          Waypoint Variable (Variable): motionParameters(jointSpeed=1.047198 jointAcceleration=1.396263 cartesianSpeed=0.09 cartesianAcceleration=0.05); variable=PSE_T_H
          URCap Gripper (Robotiq_Grippers, Robotiq Inc.) dataModel(position=24.705882352941178, force=11.0, speed=0.0, positionInDouble=24.705882352941178, forceInDouble=11.0, speedInDouble=0.0, slaveIds=[9], blocking=true)
          Waypoint Variable (Variable): variable=PSE_R
    Case (caseValue=7)
      Folder Load [hidden by the author, left out]
    Case (caseValue=8)
      Folder Unload [hidden by the author, left out]
    Case (caseValue=11)
      Folder Place without opening gripper
        Action_Info := "place object without gripper opening"
        Script: do_transition(pose_trans(FRM_Reference, PSE_T), keep_rxry=OBJ_Picked)
        Folder EXTT
          Switch expression=JIG
            Case (caseValue=1)
              Folder 3FG
                If OBJ_Picked
                  Set DigitalOutput pin=GRP_3F_Open; digitalValue=1
        If PSE_A_H≠PSE_Z
          If JNT_Q≠JNT_Z
            Script: movej(get_inverse_kin(pose_trans(FRM_Reference, PSE_A_H), qnear=JNT_Q), r=0.050)
          Else 
            Script: movej(pose_trans(FRM_Reference, PSE_A_H), r=0.050)
        If PSE_A≠PSE_Z
          If JNT_Q≠JNT_Z
            Script: movej(get_inverse_kin(pose_trans(FRM_Reference, PSE_A), qnear=JNT_Q), r=0.020)
          Else 
            Script: movej(pose_trans(FRM_Reference, PSE_A), r=0.020)
        MoveL speed 400 mm/s, acceleration 500 mm/s^2 (useActiveTCP=true) feature=FRM_Reference
          If PSE_T_H≠PSE_Z
            Waypoint Variable (Variable): motionParameters(blendRadius=0.01); variable=PSE_T_H
          Waypoint Variable (Variable): motionParameters(jointSpeed=1.047198 jointAcceleration=1.396263 cartesianSpeed=0.09 cartesianAcceleration=0.05); variable=PSE_T
            Until TOOL_CONTACT_DETECTION (allowActions=false retraction=NONE decelerationAcceleration=0.5 decelerationAngularAcceleration=34.906585)
          Force Frame feature=FRM_Reference; selection=[1, 1, 1, 0, 0, 0]; wrench=[0, 0, 0, 0, 0, 0]; limitsForce=[0.1, 0.1, 0.01, 1.047198, 1.047198, 1.047198]; limitsMotion=[0.1, 0.1, 0.1, 0.349066, 0.349066, 0.349066]
            Waypoint Variable (Variable): motionParameters(jointSpeed=1.047198 jointAcceleration=1.396263 cartesianSpeed=0.07 cartesianAcceleration=0.04); variable=PSE_T
          Folder EXTT
            Switch expression=JIG
              Case (caseValue=1)
                Folder 3FG
                  If OBJ_Picked
                    Set DigitalOutput pin=GRP_3F_Open; digitalValue=0
                    Wait Sleep waitTime=0.2
          Folder EOAT
            ''
    Case (caseValue=12)
      Folder Decap
        Action_Info := "decapping"
        Set DigitalOutput pin=GRP_3F_Enable; digitalValue=1
        Set DigitalOutput pin=GRP_3F_Decap; digitalValue=1
        Force Simple feature=Joint_6_name; selection=[0, 0, 1, 0, 0, 0]; wrench=[0, 0, 5, 0, 0, 0]; limitsForce=[0.15, 0.15, 0.15, 1.047198, 1.047198, 1.047198]; limitsMotion=[0.1, 0.1, 0.1, 0.349066, 0.349066, 0.349066]
          Script: check_decapping(offset=0.015, timeout=5, abort=CMD_Hold)
        Set DigitalOutput pin=GRP_3F_Decap; digitalValue=0
        Set DigitalOutput pin=GRP_3F_Enable; digitalValue=0
        MoveL speed 150 mm/s, acceleration 800 mm/s^2 (useActiveTCP=true) feature=FRM_Reference
          Waypoint Variable (Variable): variable=PSE_R
    Case (caseValue=13)
      Timer (action=Reset) variable(name=TMR_Barcode)
      Folder Read [hidden by the author, left out]
    Case (caseValue=15)
      Folder Detect
        Action_Info := "detect"
    Case (caseValue=30)
      Folder Shake
        Action_Info := "shake"
        Script: do_transition(pose_trans(FRM_Reference, PSE_T), keep_rxry=OBJ_Picked)
        If PSE_A_H≠PSE_Z
          If JNT_Q≠JNT_Z
            Script: movej(get_inverse_kin(pose_trans(FRM_Reference, PSE_A_H), qnear=JNT_Q), r=0.050)
          Else 
            Script: movej(pose_trans(FRM_Reference, PSE_A_H), r=0.050)
        If PSE_A≠PSE_Z
          If JNT_Q≠JNT_Z
            Script: movej(get_inverse_kin(pose_trans(FRM_Reference, PSE_A), qnear=JNT_Q), r=0.020)
          Else 
            Script: movej(pose_trans(FRM_Reference, PSE_A), r=0.020)
        MoveL speed 400 mm/s, acceleration 500 mm/s^2 (useActiveTCP=true) feature=FRM_Reference
          If PSE_T_H≠PSE_Z
            Waypoint Variable (Variable): motionParameters(blendRadius=0.01); variable=PSE_T_H
          Waypoint Variable (Variable): motionParameters(jointSpeed=1.047198 jointAcceleration=1.396263 cartesianSpeed=0.12 cartesianAcceleration=0.08); variable=PSE_T
          Folder EXTT
            ''
            MoveJ speed 60 deg/s, acceleration 80 deg/s^2 (useActiveTCP=true) feature=Base
              Waypoint Waypoint_6: TCP in base x=8.801 y=-547.927 z=402.697 mm, rx=-0.5899 ry=-0.0072 rz=-0.0613 rad; joints [-69.01, -76.872, -104.694, -56.634, 78.043, -158.781] deg; TCP offset x=0 y=0 z=161 mm, rx=3.1415 ry=0 rz=0 rad
            MoveJ speed 60 deg/s, acceleration 80 deg/s^2 (useActiveTCP=true) feature=Base
              Waypoint Waypoint_18: TCP in base x=-178.372 y=-433.927 z=368.082 mm, rx=-0.0866 ry=0.7047 rz=-0.0079 rad; joints [-72.502, -76.524, -102.817, -99.71, 50.308, -158.785] deg
            MoveJ speed 60 deg/s, acceleration 80 deg/s^2 (useActiveTCP=true) feature=Base
              Waypoint Waypoint_12: TCP in base x=8.801 y=-547.927 z=402.697 mm, rx=-0.5899 ry=-0.0072 rz=-0.0613 rad; joints [-69.01, -76.872, -104.694, -56.634, 78.043, -158.781] deg
            MoveJ speed 60 deg/s, acceleration 80 deg/s^2 (useActiveTCP=true) feature=Base
              Waypoint Waypoint_19: TCP in base x=-178.372 y=-433.927 z=368.082 mm, rx=-0.0866 ry=0.7047 rz=-0.0079 rad; joints [-72.502, -76.524, -102.817, -99.71, 50.308, -158.785] deg
          If PSE_R_H≠PSE_Z
            Waypoint Variable (Variable): motionParameters(blendRadius=0.01); variable=PSE_R
            Waypoint Variable (Variable): variable=PSE_R_H
          Else 
            Waypoint Variable (Variable): variable=PSE_R
    Case (caseValue=31)
      Action_Info := "Pick_Vial"
      Folder Pick_Vial
        URCap Gripper (Robotiq_Grippers, Robotiq Inc.) dataModel(position=0.0, force=27.84313725490196, speed=32.15686274509804, positionInDouble=0.0, forceInDouble=27.84313725490196, speedInDouble=32.15686274509804, slaveIds=[9], blocking=true)
        MoveJ speed 60 deg/s, acceleration 80 deg/s^2 (useActiveTCP=true) feature=Base
          Waypoint Vial_above: motionParameters(jointSpeed=0.436332 jointAcceleration=0.523599 cartesianSpeed=0.25 cartesianAcceleration=1.2 blendRadius=0.05); TCP in base x=17.106 y=-652.093 z=184.921 mm, rx=0 ry=0 rz=1.5641 rad; joints [-76.636, -112.403, -84.029, -73.556, 90.141, -256.27] deg
        MoveL speed 250 mm/s, acceleration 1200 mm/s^2 (useActiveTCP=true) feature=Base
          Waypoint Vial_pick_point: motionParameters(jointSpeed=1.047198 jointAcceleration=1.396263 cartesianSpeed=0.1 cartesianAcceleration=0.5); TCP in base x=17.106 y=-648.923 z=93.308 mm, rx=0 ry=0 rz=1.5641 rad; joints [-76.583, -116.742, -92.083, -61.164, 90.132, -256.177] deg
        URCap Gripper (Robotiq_Grippers, Robotiq Inc.) dataModel(position=100.0, force=32.94117647058823, speed=27.84313725490196, positionInDouble=100.0, forceInDouble=32.94117647058823, speedInDouble=27.84313725490196, slaveIds=[9], blocking=true)
        MoveL speed 250 mm/s, acceleration 1200 mm/s^2 (useActiveTCP=true) feature=Base
          Waypoint Waypoint_20: motionParameters(jointSpeed=1.047198 jointAcceleration=1.396263 cartesianSpeed=0.1 cartesianAcceleration=0.5 blendRadius=0.05); TCP in base x=19.228 y=-648.67 z=184.921 mm, rx=0 ry=0 rz=0.0241 rad; joints [-76.382, -111.96, -84.66, -73.372, 90.146, -167.779] deg
        SafeHome (positionOptionType=SPEED_AND_ACCELERATION speed=1.047198 acceleration=1.396263 nextMotionTime=2)
    Case (caseValue=32)
      decap := False
      Folder decap_Vial
        Set DigitalOutput pin=digital_out[5]; digitalValue=1
        MoveJ speed 60 deg/s, acceleration 80 deg/s^2 (useActiveTCP=true) feature=Base
          Waypoint Waypoint_47: motionParameters(jointSpeed=0.436332 jointAcceleration=0.523599 cartesianSpeed=0.25 cartesianAcceleration=1.2 blendRadius=0); TCP in base x=-32.362 y=-348.336 z=391.476 mm, rx=0 ry=0 rz=-0.0047 rad; joints [-72.819, -68.266, -97.918, -103.808, 90.124, -162.602] deg
        MoveL speed 250 mm/s, acceleration 1200 mm/s^2 (useActiveTCP=true) feature=Base
          Waypoint Vial_3FG_place: motionParameters(jointSpeed=1.047198 jointAcceleration=1.396263 cartesianSpeed=0.1 cartesianAcceleration=0.5); TCP in base x=-31.859 y=-349.403 z=145.301 mm, rx=0 ry=0 rz=0 rad; joints [-72.903, -71.756, -132.514, -65.722, 90.129, -162.805] deg
        Set DigitalOutput pin=digital_out[5]; digitalValue=0
        Wait Sleep waitTime=0.5
        MoveL speed 250 mm/s, acceleration 1200 mm/s^2 (useActiveTCP=true) feature=Base
          Waypoint Waypoint_48: motionParameters(jointSpeed=1.047198 jointAcceleration=1.396263 cartesianSpeed=0.1 cartesianAcceleration=0.5 blendRadius=0.05); TCP in base x=-32.362 y=-348.336 z=391.476 mm, rx=0 ry=0 rz=-0.0047 rad; joints [-72.819, -68.266, -97.918, -103.808, 90.124, -162.602] deg
        MoveJ speed 60 deg/s, acceleration 80 deg/s^2 (useActiveTCP=true) feature=Base
          Waypoint cap_dump: motionParameters(jointSpeed=0.436332 jointAcceleration=0.523599 cartesianSpeed=0.25 cartesianAcceleration=1.2); TCP in base x=-139.169 y=-420.164 z=146.096 mm, rx=0 ry=0 rz=0 rad; joints [-90.79, -86.479, -121, -62.513, 90.12, -180.712] deg
        URCap Gripper (Robotiq_Grippers, Robotiq Inc.) dataModel(position=0.0, force=100.0, speed=100.0, positionInDouble=0.0, forceInDouble=100.0, speedInDouble=100.0, slaveIds=[9], blocking=true)
        MoveJ speed 60 deg/s, acceleration 80 deg/s^2 (useActiveTCP=true) feature=Base
          Waypoint Waypoint_49: motionParameters(jointSpeed=0.436332 jointAcceleration=0.523599 cartesianSpeed=0.25 cartesianAcceleration=1.2 blendRadius=0.05); TCP in base x=-32.362 y=-348.336 z=391.476 mm, rx=0 ry=0 rz=-0.0047 rad; joints [-72.819, -68.266, -97.918, -103.808, 90.124, -162.602] deg
        MoveL speed 250 mm/s, acceleration 1200 mm/s^2 (useActiveTCP=true) feature=Base
          Waypoint Vial_3FG_place: motionParameters(jointSpeed=1.047198 jointAcceleration=1.396263 cartesianSpeed=0.1 cartesianAcceleration=0.5); TCP in base x=-31.859 y=-349.403 z=145.301 mm, rx=0 ry=0 rz=0 rad; joints [-72.903, -71.756, -132.514, -65.722, 90.129, -162.805] deg
        URCap Gripper (Robotiq_Grippers, Robotiq Inc.) dataModel(position=100.0, force=100.0, speed=80.0, positionInDouble=100.0, forceInDouble=100.0, speedInDouble=80.0, slaveIds=[9], blocking=true)
        SuppressedNode
          decap := True
        SuppressedNode
          Script: dynamic_upward_motion(0.015, 7)
        SuppressedNode
          MoveL speed 250 mm/s, acceleration 1200 mm/s^2 (useActiveTCP=true) feature=Joint_6_name
            MoveDirectionNode (selectedDirection=ZPlus toolParams=8.0E-4, 0.001) feature=Base
              Until DISTANCE (allowActions=false deceleration=3 distanceNodeType=STOP) Distance=0.01; motionParameters(blendRadius=0)
        SuppressedNode
          decap := False
        Folder Decap
          Action_Info := "decapping"
          Set DigitalOutput pin=GRP_3F_Enable; digitalValue=1
          Set DigitalOutput pin=GRP_3F_Decap; digitalValue=1
          Force Frame feature=Base; selection=[0, 0, 1, 0, 0, 0]; wrench=[0, 0, 1, 0, 0, 0]; limitsForce=[0.15, 0.15, 0.001, 1.047198, 1.047198, 1.047198]; limitsMotion=[0.1, 0.1, 0.1, 0.349066, 0.349066, 0.349066]
            Script: check_decapping(offset=0.015, timeout=10, abort=CMD_Hold)
          Set DigitalOutput pin=GRP_3F_Decap; digitalValue=0
          Set DigitalOutput pin=GRP_3F_Enable; digitalValue=0
          MoveL speed 250 mm/s, acceleration 1200 mm/s^2 (useActiveTCP=true) feature=Base
            Waypoint Waypoint_50: motionParameters(jointSpeed=1.047198 jointAcceleration=1.396263 cartesianSpeed=0.1 cartesianAcceleration=0.5 blendRadius=0.05); TCP in base x=-32.362 y=-348.336 z=391.476 mm, rx=0 ry=0 rz=-0.0047 rad; joints [-72.819, -68.266, -97.918, -103.808, 90.124, -162.602] deg
        MoveJ speed 60 deg/s, acceleration 80 deg/s^2 (useActiveTCP=true) feature=Base
          Waypoint cap_dump: motionParameters(jointSpeed=0.436332 jointAcceleration=0.523599 cartesianSpeed=0.25 cartesianAcceleration=1.2); TCP in base x=-139.169 y=-420.164 z=146.096 mm, rx=0 ry=0 rz=0 rad; joints [-90.79, -86.479, -121, -62.513, 90.12, -180.712] deg
        URCap Gripper (Robotiq_Grippers, Robotiq Inc.) dataModel(position=0.0, force=100.0, speed=80.0, positionInDouble=0.0, forceInDouble=100.0, speedInDouble=80.0, slaveIds=[9], blocking=true)
        MoveJ speed 60 deg/s, acceleration 80 deg/s^2 (useActiveTCP=true) feature=Base
          Waypoint Waypoint_51: motionParameters(jointSpeed=0.436332 jointAcceleration=0.523599 cartesianSpeed=0.25 cartesianAcceleration=1.2 blendRadius=0.036); TCP in base x=-32.362 y=-348.336 z=391.476 mm, rx=0 ry=0 rz=-0.0047 rad; joints [-72.819, -68.266, -97.918, -103.808, 90.124, -162.602] deg
    Case (caseValue=33)
      Folder Shake and liquid transfer
        MoveL speed 250 mm/s, acceleration 1200 mm/s^2 (useActiveTCP=true) feature=Base
          Waypoint Vial_liq_above: motionParameters(jointSpeed=1.047198 jointAcceleration=1.396263 cartesianSpeed=0.1 cartesianAcceleration=0.5); TCP in base x=-25.304 y=-338.759 z=426.628 mm, rx=-1.3159 ry=0.8 rz=-0.9283 rad; joints [-21.713, -86.8, -129.663, 45.096, -43.028, -184.708] deg
          Waypoint Vial_liq_pick_1: motionParameters(jointSpeed=1.047198 jointAcceleration=1.396263 cartesianSpeed=0.1 cartesianAcceleration=0.5); TCP in base x=-2.66 y=-335.985 z=159.39 mm, rx=-1.1505 ry=0.6732 rz=-1.0106 rad; joints [-20.975, -83.1, -137.831, -114.287, 46.064, -14.375] deg
          Waypoint Vial_liq_pick_2: motionParameters(jointSpeed=1.047198 jointAcceleration=1.396263 cartesianSpeed=0.1 cartesianAcceleration=0.5); TCP in base x=-41.402 y=-356.792 z=125.395 mm, rx=-1.1435 ry=0.6511 rz=-0.8787 rad; joints [-25.36, -82.348, -146.215, -101.788, 37.598, -24.648] deg
          URCap Gripper (Robotiq_Grippers, Robotiq Inc.) dataModel(position=100.0, force=27.84313725490196, speed=32.15686274509804, positionInDouble=100.0, forceInDouble=27.84313725490196, speedInDouble=32.15686274509804, slaveIds=[9], blocking=true)
          Wait Sleep waitTime=1
          Set DigitalOutput pin=digital_out[5]; digitalValue=1
          Wait Sleep waitTime=0.5
          Waypoint Vial_liq_above: motionParameters(jointSpeed=1.047198 jointAcceleration=1.396263 cartesianSpeed=0.05 cartesianAcceleration=0.3 blendRadius=0.05); TCP in base x=-25.304 y=-338.759 z=426.628 mm, rx=-1.3159 ry=0.8 rz=-0.9283 rad; joints [-21.713, -86.8, -129.663, 45.096, -43.028, -184.708] deg
        MoveL speed 250 mm/s, acceleration 1200 mm/s^2 (useActiveTCP=true) feature=Base
          Waypoint Liquid_midway: motionParameters(jointSpeed=1.047198 jointAcceleration=1.396263 cartesianSpeed=0.1 cartesianAcceleration=0.5 blendRadius=0); TCP in base x=57.575 y=-583.082 z=306.415 mm, rx=-1.3517 ry=0.1209 rz=-0.0969 rad; joints [-51.29, -97.606, -136.419, 36.185, 44.156, -168.768] deg
          Loop Counting (count=3) loopVariable(name=Loop_1)
            Waypoint shake_1: motionParameters(jointSpeed=1.047198 jointAcceleration=1.396263 cartesianSpeed=0.5 cartesianAcceleration=2); TCP in base x=57.575 y=-583.085 z=306.423 mm, rx=-1.361 ry=-0.1556 rz=-0.4381 rad; joints [-51.29, -97.606, -136.418, 36.185, 44.156, -145.5] deg
            Waypoint shake_2: motionParameters(jointSpeed=1.047198 jointAcceleration=1.396263 cartesianSpeed=0.5 cartesianAcceleration=2); TCP in base x=57.582 y=-583.091 z=306.44 mm, rx=-1.3088 ry=0.3685 rz=0.2149 rad; joints [-51.29, -97.606, -136.416, 36.185, 44.155, -190] deg
          Waypoint drop_above_1: motionParameters(jointSpeed=1.047198 jointAcceleration=1.396263 cartesianSpeed=0.1 cartesianAcceleration=0.5); TCP in base x=268.235 y=-467.784 z=226.22 mm, rx=-1.0278 ry=-0.4308 rz=1.0046 rad; joints [-53.609, -95.474, -138.959, 24.045, 105.829, -198.245] deg
          Waypoint drop_above_2: motionParameters(jointSpeed=1.047198 jointAcceleration=1.396263 cartesianSpeed=0.1 cartesianAcceleration=0.5); TCP in base x=219.042 y=-470.776 z=133.754 mm, rx=-0.313 ry=-0.3444 rz=1.5006 rad; joints [-60.743, -97.429, -119.175, -41.501, 111.324, -235.78] deg
          Waypoint liq_tran_1: motionParameters(jointSpeed=1.047198 jointAcceleration=1.396263 cartesianSpeed=0.05 cartesianAcceleration=0.5 blendRadius=0.008); TCP in base x=213.068 y=-469.567 z=100.231 mm, rx=0.2519 ry=0.2179 rz=1.5928 rad; joints [-44.631, -104.414, -106.819, -71.743, 78.886, -225.335] deg
          Wait Sleep waitTime=1
          Waypoint drop_above_2: motionParameters(jointSpeed=1.047198 jointAcceleration=1.396263 cartesianSpeed=0.1 cartesianAcceleration=0.5); TCP in base x=219.042 y=-470.776 z=133.754 mm, rx=-0.313 ry=-0.3444 rz=1.5006 rad; joints [-60.743, -97.429, -119.175, -41.501, 111.324, -235.78] deg
          Waypoint Waypoint_21: motionParameters(jointSpeed=1.047198 jointAcceleration=1.396263 cartesianSpeed=0.1 cartesianAcceleration=0.5); TCP in base x=187.119 y=-493.959 z=133.754 mm, rx=-0.313 ry=-0.3444 rz=1.5006 rad; joints [-65.422, -99.182, -116.519, -44.234, 112.218, -240.733] deg
          Waypoint liq_tran_2: motionParameters(jointSpeed=1.047198 jointAcceleration=1.396263 cartesianSpeed=0.05 cartesianAcceleration=0.5); TCP in base x=195.958 y=-493.023 z=100.231 mm, rx=0.1607 ry=0.1098 rz=1.5253 rad; joints [-50.52, -104.533, -106.862, -66.514, 83.832, -227.689] deg
          Wait Sleep waitTime=1
          Waypoint drop_above_2: motionParameters(jointSpeed=1.047198 jointAcceleration=1.396263 cartesianSpeed=0.1 cartesianAcceleration=0.5); TCP in base x=219.042 y=-470.776 z=133.754 mm, rx=-0.313 ry=-0.3444 rz=1.5006 rad; joints [-60.743, -97.429, -119.175, -41.501, 111.324, -235.78] deg
          Waypoint drop_above_1: motionParameters(jointSpeed=1.047198 jointAcceleration=1.396263 cartesianSpeed=0.1 cartesianAcceleration=0.5); TCP in base x=268.235 y=-467.784 z=226.22 mm, rx=-1.0278 ry=-0.4308 rz=1.0046 rad; joints [-53.609, -95.474, -138.959, 24.045, 105.829, -198.245] deg
          Waypoint Liquid_midway: motionParameters(jointSpeed=1.047198 jointAcceleration=1.396263 cartesianSpeed=0.1 cartesianAcceleration=0.5); TCP in base x=57.575 y=-583.082 z=306.415 mm, rx=-1.3517 ry=0.1209 rz=-0.0969 rad; joints [-51.29, -97.606, -136.419, 36.185, 44.156, -168.768] deg
        MoveL speed 250 mm/s, acceleration 1200 mm/s^2 (useActiveTCP=true) feature=Base
          Waypoint Vial_drop_above: motionParameters(jointSpeed=1.047198 jointAcceleration=1.396263 cartesianSpeed=0.1 cartesianAcceleration=0.5); TCP in base x=0.325 y=-648.57 z=221.894 mm, rx=-0.8735 ry=1.1659 rz=-1.4827 rad; joints [-60.601, -137.11, -52.92, -147.418, 45.283, -19.072] deg
          Waypoint Vial_liq_drop: motionParameters(jointSpeed=1.047198 jointAcceleration=1.396263 cartesianSpeed=0.1 cartesianAcceleration=0.5); TCP in base x=1.021 y=-647.66 z=92.916 mm, rx=-0.8348 ry=1.0819 rz=-1.5406 rad; joints [-60.917, -140.075, -64.676, -125.954, 46.582, -22.337] deg
          URCap Gripper (Robotiq_Grippers, Robotiq Inc.) dataModel(position=0.0, force=27.84313725490196, speed=32.15686274509804, positionInDouble=0.0, forceInDouble=27.84313725490196, speedInDouble=32.15686274509804, slaveIds=[9], blocking=true)
          Waypoint Vial_drop_above: motionParameters(jointSpeed=1.047198 jointAcceleration=1.396263 cartesianSpeed=0.1 cartesianAcceleration=0.5); TCP in base x=0.325 y=-648.57 z=221.894 mm, rx=-0.8735 ry=1.1659 rz=-1.4827 rad; joints [-60.601, -137.11, -52.92, -147.418, 45.283, -19.072] deg
    Case (caseValue=34)
      SafeHome (positionOptionType=SPEED_AND_ACCELERATION speed=1.047198 acceleration=1.396263 nextMotionTime=2)
      MoveJ speed 60 deg/s, acceleration 80 deg/s^2 (useActiveTCP=true) feature=Base
        Waypoint Waypoint_9: motionParameters(jointSpeed=0.436332 jointAcceleration=0.523599 cartesianSpeed=0.25 cartesianAcceleration=1.2); TCP in base x=206.301 y=-401.796 z=209.941 mm, rx=0 ry=0 rz=1.5608 rad; joints [-45.627, -84.145, -113.025, -72.821, 90.127, -225.014] deg
      MoveL speed 250 mm/s, acceleration 1200 mm/s^2 (useActiveTCP=true) feature=Base
        Waypoint Waypoint_10: motionParameters(jointSpeed=1.047198 jointAcceleration=1.396263 cartesianSpeed=0.1 cartesianAcceleration=0.5); TCP in base x=200.866 y=-400.818 z=105.073 mm, rx=0 ry=0 rz=1.5608 rad; joints [-46.083, -90.669, -123.933, -55.389, 90.105, -225.416] deg
      URCap Gripper (Robotiq_Grippers, Robotiq Inc.) dataModel(position=100.0, force=27.84313725490196, speed=32.15686274509804, positionInDouble=100.0, forceInDouble=27.84313725490196, speedInDouble=32.15686274509804, slaveIds=[9], blocking=true)
      Wait Sleep waitTime=1
      MoveL speed 250 mm/s, acceleration 1200 mm/s^2 (useActiveTCP=true) feature=Base
        Waypoint Waypoint_11: motionParameters(jointSpeed=1.047198 jointAcceleration=1.396263 cartesianSpeed=0.1 cartesianAcceleration=0.5 blendRadius=0.05); TCP in base x=200.866 y=-400.818 z=325.177 mm, rx=0 ry=0 rz=1.5608 rad; joints [-46.018, -81.306, -98.396, -90.289, 90.129, -225.47] deg
      MoveJ speed 60 deg/s, acceleration 80 deg/s^2 (useActiveTCP=true) feature=Base
        Waypoint Waypoint_7: motionParameters(jointSpeed=0.436332 jointAcceleration=0.523599 cartesianSpeed=0.25 cartesianAcceleration=1.2 blendRadius=0.05); TCP in base x=-615.829 y=233.809 z=300 mm, rx=0.0051 ry=0.0087 rz=-2.1118 rad; joints [-188.832, -110.936, -69.076, -89.912, 89.674, -157.919] deg
      MoveL speed 250 mm/s, acceleration 1200 mm/s^2 (useActiveTCP=true) feature=Base
        Waypoint Waypoint_8: motionParameters(jointSpeed=1.047198 jointAcceleration=1.396263 cartesianSpeed=0.1 cartesianAcceleration=0.5); TCP in base x=-615.829 y=233.809 z=13.91 mm, rx=0.0051 ry=0.0087 rz=-2.1118 rad; joints [-188.874, -123.68, -94.539, -51.707, 89.657, -157.833] deg
      URCap Gripper (Robotiq_Grippers, Robotiq Inc.) dataModel(position=0.0, force=27.84313725490196, speed=32.15686274509804, positionInDouble=0.0, forceInDouble=27.84313725490196, speedInDouble=32.15686274509804, slaveIds=[9], blocking=true)
      MoveJ speed 60 deg/s, acceleration 80 deg/s^2 (useActiveTCP=true) feature=Base
        Waypoint Waypoint_7: motionParameters(jointSpeed=0.436332 jointAcceleration=0.523599 cartesianSpeed=0.25 cartesianAcceleration=1.2); TCP in base x=-615.829 y=233.809 z=300 mm, rx=0.0051 ry=0.0087 rz=-2.1118 rad; joints [-188.832, -110.936, -69.076, -89.912, 89.674, -157.919] deg
      SafeHome (positionOptionType=SPEED_AND_ACCELERATION speed=1.047198 acceleration=1.396263 nextMotionTime=2)
      SuppressedNode
        Folder Decap
          Action_Info := "decapping"
          Set DigitalOutput pin=GRP_3F_Enable; digitalValue=1
          Set DigitalOutput pin=GRP_3F_Decap; digitalValue=1
          Force Frame feature=Base; selection=[0, 0, 1, 0, 0, 0]; wrench=[0, 0, 1, 0, 0, 0]; limitsForce=[0.15, 0.15, 0.001, 1.047198, 1.047198, 1.047198]; limitsMotion=[0.1, 0.1, 0.1, 0.349066, 0.349066, 0.349066]
            Script: check_decapping(offset=0.015, timeout=10, abort=CMD_Hold)
          Set DigitalOutput pin=GRP_3F_Decap; digitalValue=0
          Set DigitalOutput pin=GRP_3F_Enable; digitalValue=0
          MoveL speed 250 mm/s, acceleration 1200 mm/s^2 (useActiveTCP=true) feature=Base
            Waypoint Waypoint_5: motionParameters(jointSpeed=1.047198 jointAcceleration=1.396263 cartesianSpeed=0.1 cartesianAcceleration=0.5 blendRadius=0.05); TCP in base x=-31.859 y=-349.402 z=312.809 mm, rx=0 ry=0 rz=0 rad; joints [-72.832, -66.838, -110.376, -92.778, 90.139, -162.834] deg
          MoveJ speed 60 deg/s, acceleration 80 deg/s^2 (useActiveTCP=true) feature=Base
            Waypoint cap_dump: motionParameters(jointSpeed=0.436332 jointAcceleration=0.523599 cartesianSpeed=0.25 cartesianAcceleration=1.2); TCP in base x=-139.169 y=-420.164 z=146.096 mm, rx=0 ry=0 rz=0 rad; joints [-90.79, -86.479, -121, -62.513, 90.12, -180.712] deg
          URCap Gripper (Robotiq_Grippers, Robotiq Inc.) dataModel(position=0.0, force=100.0, speed=100.0, positionInDouble=0.0, forceInDouble=100.0, speedInDouble=100.0, slaveIds=[9], blocking=true)
          MoveJ speed 60 deg/s, acceleration 80 deg/s^2 (useActiveTCP=true) feature=Base
            Waypoint Waypoint_5: motionParameters(jointSpeed=0.436332 jointAcceleration=0.523599 cartesianSpeed=0.25 cartesianAcceleration=1.2 blendRadius=0.05); TCP in base x=-31.859 y=-349.402 z=312.809 mm, rx=0 ry=0 rz=0 rad; joints [-72.832, -66.838, -110.376, -92.778, 90.139, -162.834] deg
          Set DigitalOutput pin=digital_out[5]; digitalValue=1
    Case (caseValue=35)
      Folder Pick the powder container
        Wait Sleep waitTime=1
        MoveJ speed 60 deg/s, acceleration 80 deg/s^2 (useActiveTCP=true) feature=Base
          Waypoint Container_midwa: motionParameters(blendRadius=0.05); TCP in base x=-379.239 y=-127.191 z=300 mm, rx=0 ry=0 rz=-1.2472 rad; joints [-141.945, -74.312, -107.466, -88.214, 90.137, -160.485] deg
          Waypoint Container_capt: TCP in base x=-525.59 y=407.248 z=411.588 mm, rx=0 ry=0 rz=-2.8961 rad; joints [-206.083, -114.879, -46.847, -108.265, 90.132, -130.312] deg
        URCap VISOR Robotic App (SensoPart VISOR Robotic, SensoPart Industriesensorik GmbH) dataModel(visorAppTemplate=1); state(isChildrenLocked=true)
          URCap Easy Pick Setup (SensoPart VISOR Robotic, SensoPart Industriesensorik GmbH) dataModel(visorId=0, visorSetJob=true, visorJobName=Container_S, visorImageAcqSetup=2, visorCalibSetNo=7, visorDetector=1, visorImageAcqSource=0, visorOffsetSet=true, visorSetupStatus=3, Pose(key=visorImageAcqPose, Position(key=posePosition, Length(key=X value=-0.51041 unit=M), Length(key=Y value=0.417301 unit=M), Length(key=Z value=0.464095 unit=M)), Rotation(key=poseRotation, Angle(key=RX value=0.000026 unit=RAD), Angle(key=RY value=-0.000024 unit=RAD), Angle(key=RZ value=-2.896187 unit=RAD))), Pose(key=visorGripPose, Position(key=posePosition, Length(key=X value=-0.52548 unit=M), Length(key=Y value=0.459382 unit=M), Length(key=Z value=0.011872 unit=M)), Rotation(key=poseRotation, Angle(key=RX value=-0.32791 unit=RAD), Angle(key=RY value=2.076984 unit=RAD), Angle(key=RZ value=-2.068118 unit=RAD)))); state(isChildrenLocked=true)
          URCap Process (SensoPart VISOR Robotic, SensoPart Industriesensorik GmbH) dataModel(Variable(key=visorCounterVar, variable(name=easyPickCount, initializeExpression=0)), Variable(key=visorPartsFoundVar, variable(name=easyPickParts, initializeExpression=0))); state(isChildrenLocked=true)
            URCap Image Acquisition Pose (SensoPart VISOR Robotic, SensoPart Industriesensorik GmbH) state(isChildrenLocked=true)
            URCap Object Detected (SensoPart VISOR Robotic, SensoPart Industriesensorik GmbH) state(isChildrenLocked=true)
              Folder Open Gripper
                URCap Gripper (Robotiq_Grippers, Robotiq Inc.) dataModel(position=0.0, force=30.0, speed=41.84313725490196, positionInDouble=0.0, forceInDouble=30.0, speedInDouble=41.84313725490196, slaveIds=[9], blocking=true)
                MoveJ speed 60 deg/s, acceleration 80 deg/s^2 (useActiveTCP=true) feature=Base
                  Waypoint Waypoint_13: TCP in base x=-479.451 y=284.141 z=125.27 mm, rx=-0.2768 ry=2.0984 rz=-2.1213 rad; joints [-165.671, -112.009, -127.874, -95.426, 1.192, -23.029] deg
              URCap Approach Pose (SensoPart VISOR Robotic, SensoPart Industriesensorik GmbH) dataModel(visorOffsetZ=-50.0); state(isChildrenLocked=true)
              URCap Target Pose (SensoPart VISOR Robotic, SensoPart Industriesensorik GmbH) state(isChildrenLocked=true)
              Folder Close Gripper
                URCap Gripper (Robotiq_Grippers, Robotiq Inc.) dataModel(position=100.0, force=30.19607843137255, speed=41.96078431372549, positionInDouble=100.0, forceInDouble=30.19607843137255, speedInDouble=41.96078431372549, slaveIds=[9], blocking=true)
              URCap Exit Pose (SensoPart VISOR Robotic, SensoPart Industriesensorik GmbH) dataModel(visorOffsetZ=-50.0); state(isChildrenLocked=true)
            URCap No Object Detected (SensoPart VISOR Robotic, SensoPart Industriesensorik GmbH) dataModel(visorRetryCounterActive=true, Variable(key=visorNoObjCountVar, variable(name=easyPickNoObj, initializeExpression=0)))
              Popup Message (haltProgram=false message=No Container detected inputType=Text)
        MoveJ speed 60 deg/s, acceleration 80 deg/s^2 (useActiveTCP=true) feature=Base
          Waypoint Cont_midwa_1: motionParameters(blendRadius=0.05); TCP in base x=-504.067 y=246.951 z=337.123 mm, rx=-0.3472 ry=2.0343 rz=-2.0655 rad; joints [-161.564, -90.528, -130.578, -43.052, 0.855, -95.101] deg
          Waypoint Cont_midw_2: motionParameters(blendRadius=0.05); TCP in base x=-426.292 y=-118.898 z=337.123 mm, rx=-0.3472 ry=2.0343 rz=-2.0655 rad; joints [-117.656, -105.21, -94.646, -158.887, 43.73, -0.262] deg
        MoveJ speed 60 deg/s, acceleration 80 deg/s^2 (useActiveTCP=true) feature=Base
          Waypoint Waypoint_14: TCP in base x=-143.787 y=-289.021 z=255.489 mm, rx=-0.6208 ry=-1.2348 rz=1.6749 rad; joints [-116.838, -105.13, -94.648, -134.846, 121.599, 21.489] deg
          Waypoint Cont_midway_3: TCP in base x=-119.283 y=-363.048 z=317.519 mm, rx=-0.4588 ry=-0.5862 rz=1.6082 rad; joints [-109.117, -86.679, -97.632, -106.495, 122.643, 58.651] deg
          Waypoint Waypoint_43: TCP in base x=31.09 y=-542.022 z=334.788 mm, rx=-0.672 ry=-0.6244 rz=1.4088 rad; joints [-93.023, -97.009, -94.459, -77.441, 138.093, 91.25] deg
        MoveL speed 250 mm/s, acceleration 1200 mm/s^2 (useActiveTCP=true) feature=Base
          Waypoint Waypoint_27: TCP in base x=62.551 y=-565.129 z=291.796 mm, rx=-0.7505 ry=-0.749 rz=1.4123 rad; joints [-91.801, -103.314, -96.729, -71.324, 145.395, 89.047] deg
          Waypoint Waypoint_2: motionParameters(jointSpeed=1.047198 jointAcceleration=1.396263 cartesianSpeed=0.05 cartesianAcceleration=0.3); TCP in base x=-54.184 y=-562.753 z=123.32 mm, rx=-0.7505 ry=-0.749 rz=1.4123 rad; joints [-103.159, -117.824, -99.558, -69.704, 143.54, 69.763] deg
        URCap Gripper (Robotiq_Grippers, Robotiq Inc.) dataModel(position=0.0, force=100.0, speed=100.0, positionInDouble=0.0, forceInDouble=100.0, speedInDouble=100.0, slaveIds=[9], blocking=true)
        MoveL speed 250 mm/s, acceleration 1200 mm/s^2 (useActiveTCP=true) feature=Base
          Waypoint Waypoint_27: TCP in base x=62.551 y=-565.129 z=291.796 mm, rx=-0.7505 ry=-0.749 rz=1.4123 rad; joints [-91.801, -103.314, -96.729, -71.324, 145.395, 89.047] deg
          Waypoint Waypoint_39: TCP in base x=62.551 y=-565.129 z=291.796 mm, rx=-0.1058 ry=-0.0892 rz=1.5471 rad; joints [-73.149, -97.636, -88.102, -81.522, 96.755, 108.215] deg
        SafeHome (positionOptionType=SPEED_AND_ACCELERATION speed=1.047198 acceleration=1.396263 nextMotionTime=2)
        URCap VISOR Robotic App (SensoPart VISOR Robotic, SensoPart Industriesensorik GmbH) dataModel(visorAppTemplate=1); state(isChildrenLocked=true)
          URCap Easy Pick Setup (SensoPart VISOR Robotic, SensoPart Industriesensorik GmbH) dataModel(visorId=0, visorSetJob=true, visorImageAcqSetup=2, visorCalibSetNo=7, visorImageAcqSource=0, visorDetector=1, visorJobName=Target_container, visorOffsetSet=true, visorSetupStatus=4, Pose(key=visorGripPose, Position(key=posePosition, Length(key=X value=-0.64605 unit=M), Length(key=Y value=0.448738 unit=M), Length(key=Z value=0.079509 unit=M)), Rotation(key=poseRotation, Angle(key=RX value=0.000019 unit=RAD), Angle(key=RY value=-0.00001 unit=RAD), Angle(key=RZ value=-2.896171 unit=RAD))), Pose(key=visorImageAcqPose, Position(key=posePosition, Length(key=X value=-0.617993 unit=M), Length(key=Y value=0.371934 unit=M), Length(key=Z value=0.411591 unit=M)), Rotation(key=poseRotation, Angle(key=RX value=-0.000035 unit=RAD), Angle(key=RY value=-0.000001 unit=RAD), Angle(key=RZ value=-2.896152 unit=RAD)))); state(isChildrenLocked=true)
          URCap Process (SensoPart VISOR Robotic, SensoPart Industriesensorik GmbH) dataModel(Variable(key=visorCounterVar, variable(name=easyPickCount_2, initializeExpression=0)), Variable(key=visorPartsFoundVar, variable(name=easyPickParts_2, initializeExpression=0))); state(isChildrenLocked=true)
            URCap Image Acquisition Pose (SensoPart VISOR Robotic, SensoPart Industriesensorik GmbH) state(isChildrenLocked=true)
            URCap Object Detected (SensoPart VISOR Robotic, SensoPart Industriesensorik GmbH) state(isChildrenLocked=true)
              Folder Open Gripper
                URCap Gripper (Robotiq_Grippers, Robotiq Inc.) dataModel(position=0.0, force=30.0, speed=41.84313725490196, positionInDouble=0.0, forceInDouble=30.0, speedInDouble=41.84313725490196, slaveIds=[9], blocking=true)
              URCap Approach Pose (SensoPart VISOR Robotic, SensoPart Industriesensorik GmbH) dataModel(visorOffsetZ=-50.0); state(isChildrenLocked=true)
              URCap Target Pose (SensoPart VISOR Robotic, SensoPart Industriesensorik GmbH) state(isChildrenLocked=true)
              Folder Close Gripper
                URCap Gripper (Robotiq_Grippers, Robotiq Inc.) dataModel(position=100.0, force=30.19607843137255, speed=41.96078431372549, positionInDouble=100.0, forceInDouble=30.19607843137255, speedInDouble=41.96078431372549, slaveIds=[9], blocking=true)
              URCap Exit Pose (SensoPart VISOR Robotic, SensoPart Industriesensorik GmbH) dataModel(visorOffsetZ=-50.0); state(isChildrenLocked=true)
            URCap No Object Detected (SensoPart VISOR Robotic, SensoPart Industriesensorik GmbH) dataModel(visorRetryCounterActive=true, Variable(key=visorNoObjCountVar, variable(name=easyPickNoObj_2, initializeExpression=0)))
              Popup Message (haltProgram=false message=No target container is detected inputType=Text)
        MoveJ speed 60 deg/s, acceleration 80 deg/s^2 (useActiveTCP=true) feature=Base
          Waypoint Waypoint_5: TCP in base x=-545.673 y=-71.906 z=269.52 mm, rx=-0.0004 ry=-0.0002 rz=-2.9161 rad; joints [-158.416, -96.147, -92.071, -81.751, 90.145, -81.354] deg
          Waypoint Waypoint_3: TCP in base x=-19.443 y=-357.013 z=353.247 mm, rx=-0.0002 ry=-0.0003 rz=-1.8285 rad; joints [-71.157, -68.373, -103.55, -98.044, 90.131, -56.415] deg
        Set DigitalOutput pin=digital_out[5]; digitalValue=1
        MoveL speed 250 mm/s, acceleration 1200 mm/s^2 (useActiveTCP=true) feature=Base
          Waypoint Waypoint_4: TCP in base x=-27.281 y=-345.298 z=289.558 mm, rx=-0.0001 ry=-0.0003 rz=-1.2262 rad; joints [-71.854, -66.046, -114.226, -89.698, 90.15, -91.586] deg
          Waypoint Waypoint_15: motionParameters(jointSpeed=1.047198 jointAcceleration=1.396263 cartesianSpeed=0.05 cartesianAcceleration=0.3); TCP in base x=-27.267 y=-345.317 z=211.761 mm, rx=-0.0001 ry=-0.0003 rz=-1.2262 rad; joints [-71.888, -67.363, -124.926, -77.682, 90.15, -91.573] deg
        Set DigitalOutput pin=digital_out[5]; digitalValue=0
        Wait Sleep waitTime=0.5
        URCap Gripper (Robotiq_Grippers, Robotiq Inc.) dataModel(position=0.0, force=27.84313725490196, speed=49.80392156862745, positionInDouble=0.0, forceInDouble=27.84313725490196, speedInDouble=49.80392156862745, slaveIds=[9], blocking=true)
        MoveL speed 250 mm/s, acceleration 1200 mm/s^2 (useActiveTCP=true) feature=Base
          Waypoint Waypoint_16: TCP in base x=-27.285 y=-345.292 z=323.494 mm, rx=-0.0001 ry=-0.0003 rz=-1.2262 rad; joints [-71.838, -66.232, -109.162, -94.577, 90.147, -91.59] deg
        SafeHome (positionOptionType=SPEED_AND_ACCELERATION speed=1.047198 acceleration=1.396263 nextMotionTime=2)
    Case (caseValue=36)
      MoveJ speed 60 deg/s, acceleration 80 deg/s^2 (useActiveTCP=true) feature=Base
        Waypoint Waypoint_23: TCP in base x=-26.018 y=-347.731 z=350.886 mm, rx=0 ry=0 rz=-0.0073 rad; joints [-71.737, -67.031, -104.677, -98.284, 90.134, -161.343] deg
      MoveL speed 250 mm/s, acceleration 1200 mm/s^2 (useActiveTCP=true) feature=Base
        Waypoint Waypoint_24: TCP in base x=-30.861 y=-346.715 z=217.709 mm, rx=0 ry=0 rz=-0.0073 rad; joints [-72.566, -67.468, -123.973, -78.551, 90.142, -162.092] deg
      URCap Gripper (Robotiq_Grippers, Robotiq Inc.) dataModel(position=100.0, force=49.80392156862745, speed=49.80392156862745, positionInDouble=100.0, forceInDouble=49.80392156862745, speedInDouble=49.80392156862745, slaveIds=[9], blocking=true)
      Folder Decap
        Action_Info := "decapping"
        Set DigitalOutput pin=GRP_3F_Enable; digitalValue=1
        Set DigitalOutput pin=GRP_3F_Decap; digitalValue=1
        Force Frame feature=Base; selection=[0, 0, 1, 0, 0, 0]; wrench=[0, 0, 1, 0, 0, 0]; limitsForce=[0.15, 0.15, 0.001, 1.047198, 1.047198, 1.047198]; limitsMotion=[0.1, 0.1, 0.1, 0.349066, 0.349066, 0.349066]
          Script: check_decapping(offset=0.08, timeout=16, abort=CMD_Hold)
        Set DigitalOutput pin=GRP_3F_Decap; digitalValue=0
        Set DigitalOutput pin=GRP_3F_Enable; digitalValue=0
      MoveL speed 250 mm/s, acceleration 1200 mm/s^2 (useActiveTCP=true) feature=Base
        Waypoint Waypoint_17: TCP in base x=-23.963 y=-350.337 z=277.52 mm, rx=0 ry=0 rz=-0.0073 rad; joints [-71.572, -66.866, -115.515, -87.611, 90.142, -161.135] deg
        Waypoint Waypoint_22: TCP in base x=-143.535 y=-481.503 z=277.52 mm, rx=0 ry=0 rz=-0.0073 rad; joints [-91.156, -89.369, -98.021, -82.602, 90.135, -180.747] deg
        Waypoint Waypoint_25: TCP in base x=-143.535 y=-481.513 z=51.888 mm, rx=0 ry=0 rz=-0.0073 rad; joints [-91.204, -102.922, -119.604, -47.466, 90.098, -180.688] deg
      URCap Gripper (Robotiq_Grippers, Robotiq Inc.) dataModel(position=0.0, force=30.19607843137255, speed=41.96078431372549, positionInDouble=0.0, forceInDouble=30.19607843137255, speedInDouble=41.96078431372549, slaveIds=[9], blocking=true)
      MoveL speed 250 mm/s, acceleration 1200 mm/s^2 (useActiveTCP=true) feature=Base
        Waypoint Waypoint_26: TCP in base x=-143.534 y=-481.518 z=264.949 mm, rx=0 ry=0 rz=-0.0073 rad; joints [-91.159, -89.617, -99.63, -80.745, 90.135, -180.743] deg
      MoveL speed 250 mm/s, acceleration 1200 mm/s^2 (useActiveTCP=true) feature=Base
        Waypoint Waypoint_30: TCP in base x=-30.859 y=-346.719 z=243.975 mm, rx=0 ry=0 rz=-0.0073 rad; joints [-72.554, -66.791, -120.474, -82.727, 90.143, -162.097] deg
        Waypoint Waypoint_28: TCP in base x=-30.861 y=-346.715 z=174.67 mm, rx=0 ry=0 rz=-0.0073 rad; joints [-72.583, -69.344, -129.382, -71.265, 90.136, -162.084] deg
      URCap Gripper (Robotiq_Grippers, Robotiq Inc.) dataModel(position=100.0, force=30.19607843137255, speed=41.96078431372549, positionInDouble=100.0, forceInDouble=30.19607843137255, speedInDouble=41.96078431372549, slaveIds=[9], blocking=true)
      Wait Sleep waitTime=0.5
      Set DigitalOutput pin=digital_out[5]; digitalValue=1
      MoveL speed 250 mm/s, acceleration 1200 mm/s^2 (useActiveTCP=true) feature=Base
        Waypoint Waypoint_29: TCP in base x=-30.861 y=-346.715 z=297.031 mm, rx=0 ry=0 rz=-0.0073 rad; joints [-72.53, -66.334, -112.968, -90.69, 90.14, -162.104] deg
      MoveJ speed 60 deg/s, acceleration 80 deg/s^2 (useActiveTCP=true) feature=Base
        Waypoint Waypoint_31: TCP in base x=-612.104 y=16.643 z=529.968 mm, rx=0.044 ry=-0.0067 rz=-1.6589 rad; joints [-168.446, -120.76, -16.691, -134.637, 89.207, -163.626] deg
      URCap VISOR Robotic App (SensoPart VISOR Robotic, SensoPart Industriesensorik GmbH) dataModel(visorAppTemplate=1); state(isChildrenLocked=true)
        URCap Easy Pick Setup (SensoPart VISOR Robotic, SensoPart Industriesensorik GmbH) dataModel(visorId=0, visorSetJob=true, visorJobName=Weigh_scale, visorImageAcqSetup=2, visorImageAcqSource=1, visorCalibSetNo=9, visorDetector=1, visorOffsetSet=true, visorSetupStatus=2, Pose(key=visorGripPose, Position(key=posePosition, Length(key=X value=-0.680676 unit=M), Length(key=Y value=0.007363 unit=M), Length(key=Z value=0.11024 unit=M)), Rotation(key=poseRotation, Angle(key=RX value=-0.000068 unit=RAD), Angle(key=RY value=0.000005 unit=RAD), Angle(key=RZ value=-2.119482 unit=RAD)))); state(isChildrenLocked=true)
        URCap Process (SensoPart VISOR Robotic, SensoPart Industriesensorik GmbH) dataModel(Variable(key=visorCounterVar, variable(name=easyPickCount_1, initializeExpression=0)), Variable(key=visorPartsFoundVar, variable(name=easyPickParts_1, initializeExpression=0))); state(isChildrenLocked=true)
          URCap Image Acquisition Pose (SensoPart VISOR Robotic, SensoPart Industriesensorik GmbH) state(isChildrenLocked=true)
          URCap Object Detected (SensoPart VISOR Robotic, SensoPart Industriesensorik GmbH) state(isChildrenLocked=true)
            Folder Open Gripper
              Wait Sleep waitTime=0.5
            URCap Approach Pose (SensoPart VISOR Robotic, SensoPart Industriesensorik GmbH) dataModel(visorOffsetZ=-30.0); state(isChildrenLocked=true)
            URCap Target Pose (SensoPart VISOR Robotic, SensoPart Industriesensorik GmbH) state(isChildrenLocked=true)
            Folder Close Gripper
              URCap Gripper (Robotiq_Grippers, Robotiq Inc.) dataModel(position=0.0, force=100.0, speed=100.0, positionInDouble=0.0, forceInDouble=100.0, speedInDouble=100.0, slaveIds=[9], blocking=true)
            URCap Exit Pose (SensoPart VISOR Robotic, SensoPart Industriesensorik GmbH) dataModel(visorOffsetZ=-50.0); state(isChildrenLocked=true)
          URCap No Object Detected (SensoPart VISOR Robotic, SensoPart Industriesensorik GmbH) dataModel(Variable(key=visorNoObjCountVar, variable(name=easyPickNoObj_1, initializeExpression=0)))
            Popup Message (haltProgram=false message=No weigh scale detected inputType=Text)
      MoveJ speed 60 deg/s, acceleration 80 deg/s^2 (useActiveTCP=true) feature=Base
        Waypoint Waypoint_46: motionParameters(blendRadius=0.05); TCP in base x=-363.419 y=-247.513 z=293.308 mm, rx=-0.0261 ry=0.067 rz=-1.4029 rad; joints [-125.779, -78.767, -105.478, -84.647, 86.51, -135.4] deg
        Waypoint Waypoint_32: motionParameters(blendRadius=0.011); TCP in base x=49.306 y=-565.554 z=301.473 mm, rx=0.0053 ry=-0.0041 rz=-1.6935 rad; joints [-71.518, -98.113, -85.169, -86.614, 90.47, -64.53] deg
      MoveL speed 250 mm/s, acceleration 1200 mm/s^2 (useActiveTCP=true) feature=Base
        Waypoint Waypoint_33: motionParameters(blendRadius=0.05); TCP in base x=73.066 y=-562.17 z=243.824 mm, rx=-0.437 ry=0.4085 rz=-1.5974 rad; joints [-56.96, -104.117, -87.212, -96.544, 64.865, -48.999] deg
        Waypoint Waypoint_34: motionParameters(blendRadius=0.009); TCP in base x=41.968 y=-565.931 z=192.2 mm, rx=-0.4628 ry=0.4816 rz=-1.5946 rad; joints [-59.068, -107.04, -91.774, -92.086, 62.479, -49.466] deg
      URCap Gripper (Robotiq_Grippers, Robotiq Inc.) dataModel(position=79.44506104328524, force=24.19607843137255, speed=24.96078431372549, positionInDouble=79.44506104328524, forceInDouble=24.19607843137255, speedInDouble=24.96078431372549, slaveIds=[9], blocking=true)
      MoveL speed 250 mm/s, acceleration 1200 mm/s^2 (useActiveTCP=true) feature=Base
        Waypoint Waypoint_40: motionParameters(blendRadius=0.001); TCP in base x=42.988 y=-565.986 z=193.701 mm, rx=-0.0174 ry=0.5963 rz=-0.1501 rad; joints [-58.912, -106.823, -91.879, -91.953, 62.347, -134.939] deg
        Waypoint decap_1: motionParameters(blendRadius=0); TCP in base x=44.392 y=-566.054 z=195.773 mm, rx=0.7594 ry=0.2073 rz=2.4462 rad; joints [-58.665, -106.535, -92.031, -91.804, 62.093, -289.256] deg
      URCap Gripper (Robotiq_Grippers, Robotiq Inc.) dataModel(position=15.738068812430626, force=60.0, speed=67.84313725490196, positionInDouble=15.738068812430626, forceInDouble=60.0, speedInDouble=67.84313725490196, slaveIds=[9], blocking=true)
      MoveL speed 250 mm/s, acceleration 1200 mm/s^2 (useActiveTCP=true) feature=Base
        Waypoint Waypoint_41: motionParameters(blendRadius=0); TCP in base x=44.392 y=-566.054 z=195.773 mm, rx=0.4124 ry=0.4915 rz=1.2883 rad; joints [-58.667, -106.534, -92.032, -91.801, 62.096, -219.81] deg
        Waypoint Waypoint_42: motionParameters(blendRadius=0); TCP in base x=44.392 y=-566.054 z=195.773 mm, rx=-0.2725 ry=0.5572 rz=-0.9456 rad; joints [-58.67, -106.534, -92.029, -91.8, 62.103, -87.689] deg
        Waypoint decap_2: motionParameters(blendRadius=0); TCP in base x=44.392 y=-566.054 z=195.773 mm, rx=0.8954 ry=0.0162 rz=2.9091 rad; joints [-58.667, -106.534, -92.032, -91.801, 62.096, 42.276] deg; TCP offset x=0 y=0 z=161 mm, rx=3.1415 ry=0 rz=0 rad
      URCap Gripper (Robotiq_Grippers, Robotiq Inc.) dataModel(position=79.44506104328524, force=31.0, speed=38.84313725490196, positionInDouble=79.44506104328524, forceInDouble=31.0, speedInDouble=38.84313725490196, slaveIds=[9], blocking=true)
      MoveL speed 250 mm/s, acceleration 1200 mm/s^2 (useActiveTCP=true) feature=Base
        Waypoint Waypoint_44: motionParameters(blendRadius=0); TCP in base x=44.392 y=-566.054 z=195.773 mm, rx=-0.419 ry=0.4993 rz=-1.4153 rad; joints [-58.666, -106.534, -92.032, -91.802, 62.095, -59.805] deg; TCP offset x=0 y=0 z=161 mm, rx=3.1415 ry=0 rz=0 rad
        Waypoint Waypoint_45: motionParameters(blendRadius=0); TCP in base x=44.392 y=-566.054 z=195.773 mm, rx=0.1471 ry=0.5829 rz=0.4157 rad; joints [-58.664, -106.539, -92.027, -91.813, 62.089, -168.131] deg
        Waypoint decap_1: motionParameters(blendRadius=0); TCP in base x=44.392 y=-566.054 z=195.773 mm, rx=0.7594 ry=0.2073 rz=2.4462 rad; joints [-58.665, -106.535, -92.031, -91.804, 62.093, -289.256] deg
        Waypoint Waypoint_35: motionParameters(blendRadius=0); TCP in base x=80.306 y=-567.231 z=248.688 mm, rx=0.7594 ry=0.2073 rz=2.4462 rad; joints [-55.796, -106.6, -83.626, -101.521, 63.116, -286.278] deg
        Waypoint Waypoint_36: motionParameters(blendRadius=0); TCP in base x=80.289 y=-567.231 z=248.695 mm, rx=0 ry=0 rz=2.4462 rad; joints [-68.422, -99.693, -91.068, -79.223, 90.134, -298.595] deg
        Waypoint Waypoint_37: motionParameters(blendRadius=0.05); TCP in base x=-160.607 y=-659.592 z=248.695 mm, rx=0 ry=0 rz=2.4462 rad; joints [-92.274, -114.356, -71.715, -83.911, 90.147, -322.496] deg
        Waypoint Waypoint_38: motionParameters(blendRadius=0.05); TCP in base x=-156.656 y=-635.547 z=54.757 mm, rx=0 ry=0 rz=2.4462 rad; joints [-92.043, -120.062, -93.338, -56.583, 90.13, -322.166] deg
      URCap Gripper (Robotiq_Grippers, Robotiq Inc.) dataModel(position=28.479467258601545, force=60.0, speed=67.84313725490196, positionInDouble=28.479467258601545, forceInDouble=60.0, speedInDouble=67.84313725490196, slaveIds=[9], blocking=true)
      MoveL speed 250 mm/s, acceleration 1200 mm/s^2 (useActiveTCP=true) feature=Base
        Waypoint Waypoint_37: motionParameters(blendRadius=0.05); TCP in base x=-160.607 y=-659.592 z=248.695 mm, rx=0 ry=0 rz=2.4462 rad; joints [-92.274, -114.356, -71.715, -83.911, 90.147, -322.496] deg
      SafeHome (positionOptionType=SPEED_AND_ACCELERATION speed=1.047198 acceleration=1.396263 nextMotionTime=2)
    Case (caseValue=37)
      Folder Detect spatula and powder transfer
        URCap VISOR Robotic App (SensoPart VISOR Robotic, SensoPart Industriesensorik GmbH) dataModel(visorAppTemplate=1); state(isChildrenLocked=true)
          URCap Easy Pick Setup (SensoPart VISOR Robotic, SensoPart Industriesensorik GmbH) dataModel(visorId=0, visorSetJob=true, visorJobName=Spatula, visorImageAcqSetup=2, visorImageAcqSource=1, visorCalibSetNo=10, visorDetector=1, visorOffsetSet=true, visorSetupStatus=2, Pose(key=visorGripPose, Position(key=posePosition, Length(key=X value=-0.66033 unit=M), Length(key=Y value=-0.361002 unit=M), Length(key=Z value=0.13373 unit=M)), Rotation(key=poseRotation, Angle(key=RX value=-0.000075 unit=RAD), Angle(key=RY value=-0.000089 unit=RAD), Angle(key=RZ value=-0.086276 unit=RAD)))); state(isChildrenLocked=true)
          URCap Process (SensoPart VISOR Robotic, SensoPart Industriesensorik GmbH) dataModel(Variable(key=visorCounterVar, variable(name=easyPickCount_3, initializeExpression=0)), Variable(key=visorPartsFoundVar, variable(name=easyPickParts_3, initializeExpression=0))); state(isChildrenLocked=true)
            URCap Image Acquisition Pose (SensoPart VISOR Robotic, SensoPart Industriesensorik GmbH) state(isChildrenLocked=true)
            URCap Object Detected (SensoPart VISOR Robotic, SensoPart Industriesensorik GmbH) state(isChildrenLocked=true)
              Folder Open Gripper
                URCap Gripper (Robotiq_Grippers, Robotiq Inc.) dataModel(position=0.0, force=34.90196078431372, speed=50.98039215686274, positionInDouble=0.0, forceInDouble=34.90196078431372, speedInDouble=50.98039215686274, slaveIds=[9], blocking=true)
              URCap Approach Pose (SensoPart VISOR Robotic, SensoPart Industriesensorik GmbH) dataModel(visorOffsetZ=-100.0); state(isChildrenLocked=true)
              URCap Target Pose (SensoPart VISOR Robotic, SensoPart Industriesensorik GmbH) state(isChildrenLocked=true)
              Folder Close Gripper
                URCap Gripper (Robotiq_Grippers, Robotiq Inc.) dataModel(position=100.0, force=35.0, speed=51.0, positionInDouble=100.0, forceInDouble=35.0, speedInDouble=51.0, slaveIds=[9], blocking=true)
              URCap Exit Pose (SensoPart VISOR Robotic, SensoPart Industriesensorik GmbH) dataModel(visorOffsetZ=-200.0); state(isChildrenLocked=true)
            URCap No Object Detected (SensoPart VISOR Robotic, SensoPart Industriesensorik GmbH) dataModel(Variable(key=visorNoObjCountVar, variable(name=easyPickNoObj_3, initializeExpression=0)))
              Popup Message (haltProgram=false message=No spatula is detected inputType=Text)
        MoveL speed 250 mm/s, acceleration 1200 mm/s^2 (useActiveTCP=true) feature=Base
          Waypoint Waypoint_52: TCP in base x=-311.184 y=-360.981 z=333.55 mm, rx=-0.0353 ry=0.8169 rz=-0.0814 rad; joints [-88.031, -71.899, -115.722, -84.491, 43.339, 187.849] deg
          Waypoint Waypoint_53: motionParameters(jointSpeed=1.047198 jointAcceleration=1.396263 cartesianSpeed=0.05 cartesianAcceleration=0.3); TCP in base x=205.605 y=-570.795 z=367.492 mm, rx=-0.0353 ry=0.8169 rz=-0.0814 rad; joints [-44.083, -120.726, -47.91, -138.679, 59.535, 241.172] deg
          Loop Counting (count=2) loopVariable(name=Loop_2)
            Waypoint Waypoint_54: motionParameters(jointSpeed=1.047198 jointAcceleration=1.396263 cartesianSpeed=0.05 cartesianAcceleration=0.3); TCP in base x=82.882 y=-561.436 z=212.22 mm, rx=-0.0362 ry=0.7929 rz=-0.0809 rad; joints [-51.957, -110.229, -86.761, -104.901, 55.879, 232.906] deg
              Until TOOL_CONTACT_DETECTION (allowActions=false retraction=0 decelerationAcceleration=3 decelerationAngularAcceleration=34.906585)
            Waypoint Waypoint_55: motionParameters(jointSpeed=1.047198 jointAcceleration=1.396263 cartesianSpeed=0.05 cartesianAcceleration=0.3); TCP in base x=114.847 y=-565.201 z=237.656 mm, rx=-0.0274 ry=1.0163 rz=-0.0859 rad; joints [-47.723, -117.859, -75.471, -124.529, 51.946, 244.966] deg
            Waypoint Waypoint_56: motionParameters(jointSpeed=1.047198 jointAcceleration=1.396263 cartesianSpeed=0.05 cartesianAcceleration=0.3); TCP in base x=154.686 y=-566.893 z=248.204 mm, rx=-0.0235 ry=1.1118 rz=-0.0878 rad; joints [-44.701, -123.843, -66.489, -135.419, 52.27, 251.271] deg
          Waypoint Waypoint_57: motionParameters(jointSpeed=1.047198 jointAcceleration=1.396263 cartesianSpeed=0.75 cartesianAcceleration=1.5); TCP in base x=154.686 y=-566.893 z=230.068 mm, rx=-0.0235 ry=1.1118 rz=-0.0878 rad; joints [-44.704, -124.369, -68.338, -133.046, 52.276, 251.276] deg
          Waypoint Waypoint_56: motionParameters(jointSpeed=1.047198 jointAcceleration=1.396263 cartesianSpeed=0.05 cartesianAcceleration=0.3 blendRadius=0.017); TCP in base x=154.686 y=-566.893 z=248.204 mm, rx=-0.0235 ry=1.1118 rz=-0.0878 rad; joints [-44.701, -123.843, -66.489, -135.419, 52.27, 251.271] deg
          Waypoint Waypoint_58: motionParameters(jointSpeed=1.047198 jointAcceleration=1.396263 cartesianSpeed=0.05 cartesianAcceleration=0.3 blendRadius=0.05); TCP in base x=231.567 y=-569.526 z=278.594 mm, rx=0.0007 ry=1.6481 rz=-0.0969 rad; joints [-39.887, -150.285, -32.053, -182.923, 53.747, 276.565] deg
          Waypoint Waypoint_59: motionParameters(jointSpeed=1.047198 jointAcceleration=1.396263 cartesianSpeed=0.05 cartesianAcceleration=0.3 blendRadius=0.05); TCP in base x=1.876 y=-569.571 z=422.253 mm, rx=-0.0127 ry=1.6478 rz=-0.0845 rad; joints [-53.633, -124.815, -56.782, -185.119, 39.184, 278.728] deg
          Waypoint Waypoint_60: motionParameters(blendRadius=0.05); TCP in base x=-440.228 y=-361.405 z=422.253 mm, rx=0.7186 ry=1.5438 rz=-0.7545 rad; joints [-104.438, -124.815, -56.782, -185.119, 39.184, 278.728] deg
          Waypoint Waypoint_61: motionParameters(blendRadius=0.05); TCP in base x=-538.505 y=-132.796 z=241.168 mm, rx=0.6097 ry=1.5298 rz=-0.6765 rad; joints [-122.081, -111.603, -103.756, -151.61, 14.953, 280.114] deg
          Waypoint Waypoint_62: TCP in base x=-541.29 y=-135.432 z=161.029 mm, rx=0.6351 ry=1.5212 rz=-0.7033 rad; joints [-122.481, -119.984, -105.433, -140.609, 16.478, 279.223] deg
          Waypoint Waypoint_63: motionParameters(jointSpeed=1.047198 jointAcceleration=1.396263 cartesianSpeed=0.02 cartesianAcceleration=0.1); TCP in base x=-584.28 y=-74.564 z=291.281 mm, rx=0.2441 ry=0.6849 rz=-0.8345 rad; joints [-141.987, -91.134, -105.079, -67.56, 50.134, 175.736] deg
            SuppressedNode
              Until EXPRESSION (allowActions=false) ExpressionBranch=Weight_value<32
        SuppressedNode
          Loop While (checkContinuously=true) expression=Weight_value>32.000
            MoveL speed 250 mm/s, acceleration 1200 mm/s^2 (useActiveTCP=true) feature=Base
              Waypoint Waypoint_52: motionParameters(blendRadius=0.05); TCP in base x=-311.184 y=-360.981 z=333.55 mm, rx=-0.0353 ry=0.8169 rz=-0.0814 rad; joints [-88.031, -71.899, -115.722, -84.491, 43.339, 187.849] deg
              Waypoint Waypoint_53: motionParameters(jointSpeed=1.047198 jointAcceleration=1.396263 cartesianSpeed=0.05 cartesianAcceleration=0.3); TCP in base x=205.605 y=-570.795 z=367.492 mm, rx=-0.0353 ry=0.8169 rz=-0.0814 rad; joints [-44.083, -120.726, -47.91, -138.679, 59.535, 241.172] deg
              Loop Counting (count=2) loopVariable(name=Loop_5)
                Waypoint Waypoint_54: motionParameters(jointSpeed=1.047198 jointAcceleration=1.396263 cartesianSpeed=0.05 cartesianAcceleration=0.3); TCP in base x=82.882 y=-561.436 z=212.22 mm, rx=-0.0362 ry=0.7929 rz=-0.0809 rad; joints [-51.957, -110.229, -86.761, -104.901, 55.879, 232.906] deg
                  Until TOOL_CONTACT_DETECTION (allowActions=false retraction=0 decelerationAcceleration=3 decelerationAngularAcceleration=34.906585)
                Waypoint Waypoint_55: motionParameters(jointSpeed=1.047198 jointAcceleration=1.396263 cartesianSpeed=0.05 cartesianAcceleration=0.3); TCP in base x=114.847 y=-565.201 z=237.656 mm, rx=-0.0274 ry=1.0163 rz=-0.0859 rad; joints [-47.723, -117.859, -75.471, -124.529, 51.946, 244.966] deg
                Waypoint Waypoint_56: motionParameters(jointSpeed=1.047198 jointAcceleration=1.396263 cartesianSpeed=0.05 cartesianAcceleration=0.3); TCP in base x=154.686 y=-566.893 z=248.204 mm, rx=-0.0235 ry=1.1118 rz=-0.0878 rad; joints [-44.701, -123.843, -66.489, -135.419, 52.27, 251.271] deg
              Waypoint Waypoint_57: motionParameters(jointSpeed=1.047198 jointAcceleration=1.396263 cartesianSpeed=0.75 cartesianAcceleration=1.5); TCP in base x=154.686 y=-566.893 z=230.068 mm, rx=-0.0235 ry=1.1118 rz=-0.0878 rad; joints [-44.704, -124.369, -68.338, -133.046, 52.276, 251.276] deg
              Waypoint Waypoint_56: motionParameters(jointSpeed=1.047198 jointAcceleration=1.396263 cartesianSpeed=0.05 cartesianAcceleration=0.3 blendRadius=0.017); TCP in base x=154.686 y=-566.893 z=248.204 mm, rx=-0.0235 ry=1.1118 rz=-0.0878 rad; joints [-44.701, -123.843, -66.489, -135.419, 52.27, 251.271] deg
              Waypoint Waypoint_58: motionParameters(jointSpeed=1.047198 jointAcceleration=1.396263 cartesianSpeed=0.05 cartesianAcceleration=0.3 blendRadius=0.05); TCP in base x=231.567 y=-569.526 z=278.594 mm, rx=0.0007 ry=1.6481 rz=-0.0969 rad; joints [-39.887, -150.285, -32.053, -182.923, 53.747, 276.565] deg
              Waypoint Waypoint_59: motionParameters(jointSpeed=1.047198 jointAcceleration=1.396263 cartesianSpeed=0.05 cartesianAcceleration=0.3 blendRadius=0.05); TCP in base x=1.876 y=-569.571 z=422.253 mm, rx=-0.0127 ry=1.6478 rz=-0.0845 rad; joints [-53.633, -124.815, -56.782, -185.119, 39.184, 278.728] deg
              Waypoint Waypoint_60: motionParameters(blendRadius=0.05); TCP in base x=-440.228 y=-361.405 z=422.253 mm, rx=0.7186 ry=1.5438 rz=-0.7545 rad; joints [-104.438, -124.815, -56.782, -185.119, 39.184, 278.728] deg
              Waypoint Waypoint_61: motionParameters(blendRadius=0.05); TCP in base x=-538.505 y=-132.796 z=241.168 mm, rx=0.6097 ry=1.5298 rz=-0.6765 rad; joints [-122.081, -111.603, -103.756, -151.61, 14.953, 280.114] deg
              Waypoint Waypoint_62: TCP in base x=-541.29 y=-135.432 z=161.029 mm, rx=0.6351 ry=1.5212 rz=-0.7033 rad; joints [-122.481, -119.984, -105.433, -140.609, 16.478, 279.223] deg
              Waypoint Waypoint_63: motionParameters(jointSpeed=1.047198 jointAcceleration=1.396263 cartesianSpeed=0.02 cartesianAcceleration=0.1); TCP in base x=-584.28 y=-74.564 z=291.281 mm, rx=0.2441 ry=0.6849 rz=-0.8345 rad; joints [-141.987, -91.134, -105.079, -67.56, 50.134, 175.736] deg
  '=========='
  Folder PostSettings [hidden by the author, left out]
